# B&R Automation Studio project BoostTest
Automation Studio 6.7.2.9; technology packages: OpcUaCs 6.0.0

## Configuration CgAutomation

CPU X20EM0611, AutomationRuntime 6.3.4, Build 11.3.0, Vc 6.0.0

### Task classes (Cpu.sw)
```
Cyclic#1:
  Prg01 <- Machine.Prg01.prg
Cyclic#2:
  Prg02 <- Machine.Prg02.prg
Binaries: udbdef, FWRules, TCData, sysconf, iomap, ashwd, BRRole, asfw, arconfig, ashwac, UaCsConfig
Libraries: sys_lib, runtime, CFrw, CAlarm, astime, AsIecCon, CPrg01, CPrg02
```

### Hardware
```
X20EM0611 : X20EM0611 v1.1.1.0
  Connector IF2:
    ActivateDevice = 1
  ConfigurationID = BoostTest_CgAutomation
  Simulation = 1
  FileDevice1
  FileDeviceName1 = USER
  FileDevicePath1 = USER_PATH
```

### BRRole.brrole - X20EM0611/AccessAndSecurity/UserRoleSystem/BRRole.brrole
```
Element BR_Anonymous (Type=BRRole)
Element BR_Engineer (Type=BRRole)
Element BR_Observer (Type=BRRole)
Element BR_SafetyAdmin (Type=BRRole)
Element BR_SecurityAdmin (Type=BRRole)
```

- Safety project (password-protected, skipped)

## Logical view

Binary libraries used (declarations not repeated): operator, runtime, AsIecCon, astime, sys_lib

### Package Logical/Libraries - Global libraries

### Framework.st
```iecst
ACTION aFrwInit:
	ST_name(0, ADR(sObjName), 0);
END_ACTION

ACTION aFrwCyclic:

	aPreStateExt;
	aCallRessource;
	CASE stModuleData.enModuleState OF

		enState_Initialising:
            aInitialisingExt;
            IF (stModuleData.bInitDone) THEN
                stModuleData.enModuleState := enState_Stopped;
            END_IF

		enState_Stopped:
			aStoppedExt;

		enState_Running:
			aRunningExt;

		ELSE
			stModuleData.enModuleState := enState_Initialising;
	END_CASE

	aPostStateExt;

END_ACTION

ACTION aRessource_01:
    udiRessource_01 := udiRessource_01 + 1;
END_ACTION

ACTION aRessource_02:
    udiRessource_02 := udiRessource_02 + 2;
END_ACTION
```

### Framework.var
```iecst
VAR
    _ii : INT;
    sObjName : STRING[10];
    dstAlarm : REFERENCE TO tstCFrw_AlarmType;
END_VAR
(*Sub-States*)
VAR
    stInitialisingExt : tstInitialisingExt;
    stRunExt : tstRunExt;
    New_Variable : USINT;
END_VAR
```

### Library Logical/Framework/Ressources/CFrw (IEC)

#### Types.typ - Exported data types
```iecst
TYPE
	tenCFrw_States :
		(
		enState_Initialising,
		enState_Stopped,
		enState_Running
		);
	tstCFrw_AlarmType : 	STRUCT
		sDefaultText : STRING[255];
		udiCode : UDINT;
		uiSeverity : UINT;
	END_STRUCT;
END_TYPE
```

### Ressource_01.var
```iecst
VAR
    udiRessource_01 : UDINT;
END_VAR
```

### Ressource_01.st
```iecst
ACTION aCallRessource:
    aRessource_01;
    aReferencedAction;
END_ACTION

ACTION aReferencedAction:
    aLocalAction;
END_ACTION
```

### Ressource_02.var
```iecst
VAR
    udiRessource_02 : UDINT;
END_VAR
```

### Ressource_02.st
```iecst
ACTION aCallRessource:
    aRessource_02;
END_ACTION
```

### Program Logical/Framework/Template/Template (IEC)

- Framework.st (reference to Logical/Framework/Ressources/Framework.st)

- Framework.var (reference to Logical/Framework/Ressources/Framework.var)

#### Cyclic.st - Cyclic code
```iecst
PROGRAM _CYCLIC
	(* Insert code here *)
	 aFrwCyclic;
END_PROGRAM
```

#### Init.st - Init code
```iecst
PROGRAM _INIT
	(* Insert code here *)
	aFrwInit;

END_PROGRAM
```

#### Exit.st - Exit code
```iecst
PROGRAM _EXIT
	(* Insert code here *)

END_PROGRAM
```

#### Template.typ - Local data types
```iecst
TYPE
    tstAlarmList :     STRUCT
        stFrwAlarms : tstCAlarm_FrwAlarmListType;
        stModuleAlarms : tst_TEMPL_AlarmType;
    END_STRUCT;
    tst_TEMPL_AlarmType :     STRUCT
        stAlarm500000 : tstAlarm500000;
    END_STRUCT;
END_TYPE

(*States*)

TYPE
    tstInitialisingExt :     STRUCT
        enState : tenInitialisingExt;
    END_STRUCT;
    tenInitialisingExt :
        (
        enInitialisingExt_EntryAction,
        enInitialisingExt_, (*insert machine specific states here*)
        enInitialisingExt_Done
        );
    tstRunExt :     STRUCT
        enState : tenRunExt;
    END_STRUCT;
    tenRunExt :
        (
        enRunExt_EntryAction,
        enRunExt_, (*insert machine specific states here*)
        enRunExt_Done
        );
END_TYPE
```

#### Template.var - Local variables
```iecst
VAR
    stAlarmList : tstAlarmList;
    stModuleData : tstC_TEMPL_Data;
END_VAR
```

#### PreStateExt.st
```iecst
ACTION aPreStateExt:

END_ACTION
```

#### States.st
```iecst
ACTION aInitialisingExt:
    CASE stInitialisingExt.enState OF
        enInitialisingExt_EntryAction:
            stInitialisingExt.enState := enInitialisingExt_;
        enInitialisingExt_:
            (*implement machine specific code here*)
            stInitialisingExt.enState := enInitialisingExt_Done;
        enInitialisingExt_Done:
            (*set bInitDone := TRUE if initialising is completed*)
            stModuleData.bInitDone := TRUE;
        ELSE
            ;
    END_CASE
END_ACTION

ACTION aStoppedExt:

END_ACTION

ACTION aRunningExt:

END_ACTION
```

#### PostStateExt.st
```iecst
ACTION aPostStateExt:

END_ACTION
```

### Library Logical/Framework/Template/C_TEMPL_ (IEC)

#### C_TEMPL_.typ - Exported data types
```iecst
TYPE
    tstC_TEMPL_Data :     STRUCT
        enModuleState : tenCFrw_States;
        bInitDone : BOOL;
        stPar : tstC_TEMPL_Par;
    END_STRUCT;
    tstC_TEMPL_Par :     STRUCT
        udiPar01 : UDINT;
    END_STRUCT;
END_TYPE
```

### Library Logical/Machine/CAlarm (IEC)

#### Types.typ - Exported data types
```iecst
(*Framework*)

TYPE
	tstAlarm100000 :tstCFrw_AlarmType := (sDefaultText:='Message 100000',udiCode:=100000);
	tstAlarm100001 :tstCFrw_AlarmType := (sDefaultText:='Message 100001',udiCode:=100001);
	tstAlarm100002 :tstCFrw_AlarmType := (sDefaultText:='Message 100002',udiCode:=100002);
	tstCAlarm_FrwAlarmListType : 	STRUCT
		stAlarm100000 : tstAlarm100000;
		stAlarm100001 : tstAlarm100001;
		stAlarm100002 : tstAlarm100002;
	END_STRUCT;
END_TYPE

(*Process*)

TYPE
	tstAlarm500000 :tstCFrw_AlarmType := (sDefaultText:='Message 500000',udiCode:=500000);
	tstAlarm500001 :tstCFrw_AlarmType := (sDefaultText:='Message 500001',udiCode:=500001);
END_TYPE
```

### Program Logical/Machine/Prg01 (IEC)

- Framework.st (reference to Logical/Framework/Ressources/Framework.st)

- Framework.var (reference to Logical/Framework/Ressources/Framework.var)

- Ressource_01.var (reference to Logical/Framework/Ressources/Ressource_01/Ressource_01.var)

- Ressource_01.st (reference to Logical/Framework/Ressources/Ressource_01/Ressource_01.st)

#### Action.st
```iecst
ACTION aLocalAction:
    sText := 'aLocalAction called';
END_ACTION
```

#### Cyclic.st - Cyclic code
```iecst
PROGRAM _CYCLIC
	(* Insert code here *)
    aFrwCyclic;
    udiRessource_01;
END_PROGRAM
```

#### Init.st - Init code
```iecst
PROGRAM _INIT
	(* Insert code here *)
	aFrwInit;

END_PROGRAM
```

#### Exit.st - Exit code
```iecst
PROGRAM _EXIT
	(* Insert code here *)

END_PROGRAM
```

#### Prg01.typ - Local data types
```iecst
TYPE
    tstAlarmList :     STRUCT
        stFrwAlarms : tstCAlarm_FrwAlarmListType;
        stModuleAlarms : tstPrg01_AlarmType;
    END_STRUCT;
    tstPrg01_AlarmType :     STRUCT
        stAlarm500000 : tstAlarm500000;
    END_STRUCT;
END_TYPE

(*States*)

TYPE
    tstInitialisingExt :     STRUCT
        enState : tenInitialisingExt;
    END_STRUCT;
    tenInitialisingExt :
        (
        enInitialisingExt_EntryAction,
        enInitialisingExt_InitPrg01, (*insert machine specific states here*)
        enInitialisingExt_Done
        );
    tstRunExt :     STRUCT
        enState : tenRunExt;
    END_STRUCT;
    tenRunExt :
        (
        enRunExt_EntryAction,
        enRunExt_, (*insert machine specific states here*)
        enRunExt_Done
        );
    tstDebugStruct :     STRUCT
        bFlag : BOOL;
        diValue : DINT;
    END_STRUCT;
END_TYPE
```

#### Prg01.var - Local variables
```iecst
VAR
    stAlarmList : tstAlarmList;
    stModuleData : tstCPrg01Data;
    sText : STRING[80];
    pDebugArray : UDINT;
    astDebugArray : ARRAY[0..1] OF tstDebugStruct;
    dastDebugArray : REFERENCE TO ARRAY[0..1] OF tstDebugStruct;
END_VAR
```

#### PreStateExt.st
```iecst
ACTION aPreStateExt:
    pDebugArray := ADR(astDebugArray);
    dastDebugArray ACCESS pDebugArray;
END_ACTION
```

#### States.st
```iecst
ACTION aInitialisingExt:

    CASE stInitialisingExt.enState OF
        enInitialisingExt_EntryAction:
            stInitialisingExt.enState := enInitialisingExt_InitPrg01;
        enInitialisingExt_InitPrg01:
            (*implement machine specific code here*)
            stInitialisingExt.enState := enInitialisingExt_Done;
        enInitialisingExt_Done:
            (*set bInitDone := TRUE if initialising is completed*)
            stModuleData.bInitDone := TRUE;
        ELSE
            ;
    END_CASE
END_ACTION

ACTION aStoppedExt:

	FOR _ii := 0 TO 5 DO
		;
	END_FOR

END_ACTION

ACTION aRunningExt:

END_ACTION
```

#### PostStateExt.st
```iecst
ACTION aPostStateExt:

	FOR _ii := 0 TO (SIZEOF(stAlarmList.stFrwAlarms)/SIZEOF(dstAlarm) - 1) DO
		dstAlarm ACCESS ADR(stAlarmList.stFrwAlarms) + _ii * SIZEOF(dstAlarm);
	END_FOR

END_ACTION
```

### Library Logical/Machine/CPrg01 (IEC)

#### CPrg01.typ - Exported data types
```iecst
TYPE
    tstCPrg01Data :     STRUCT
        enModuleState : tenCFrw_States;
        bInitDone : BOOL;
        stPar : tstCPrg01Par;
    END_STRUCT;
    tstCPrg01Par :     STRUCT
        udiPar01 : UDINT;
    END_STRUCT;
END_TYPE
```

### Program Logical/Machine/Prg02 (IEC)

- Framework.st (reference to Logical/Framework/Ressources/Framework.st)

- Framework.var (reference to Logical/Framework/Ressources/Framework.var)

- Ressource_02.var (reference to Logical/Framework/Ressources/Ressource_02/Ressource_02.var)

- Ressource_02.st (reference to Logical/Framework/Ressources/Ressource_02/Ressource_02.st)

#### Cyclic.st - Cyclic code
```iecst
PROGRAM _CYCLIC
	(* Insert code here *)
    aFrwCyclic;
    udiRessource_02;
END_PROGRAM
```

#### Init.st - Init code
```iecst
PROGRAM _INIT
	(* Insert code here *)
	aFrwInit;

END_PROGRAM
```

#### Exit.st - Exit code
```iecst
PROGRAM _EXIT
	(* Insert code here *)

END_PROGRAM
```

#### Prg02.typ - Local data types
```iecst
TYPE
    tstAlarmList :     STRUCT
        stFrwAlarms : tstCAlarm_FrwAlarmListType;
        stModuleAlarms : tstPrg02_AlarmType;
    END_STRUCT;
    tstPrg02_AlarmType :     STRUCT
        stAlarm500001 : tstAlarm500001;
    END_STRUCT;
END_TYPE

(*States*)

TYPE
    tstInitialisingExt :     STRUCT
        enState : tenInitialisingExt;
    END_STRUCT;
    tenInitialisingExt :
        (
        enInitialisingExt_EntryAction,
        enInitialisingExt_InitPrg02, (*insert machine specific states here*)
        enInitialisingExt_Done
        );
    tstRunExt :     STRUCT
        enState : tenRunExt;
    END_STRUCT;
    tenRunExt :
        (
        enRunExt_EntryAction,
        enRunExt_, (*insert machine specific states here*)
        enRunExt_Done
        );
END_TYPE
```

#### Prg02.var - Local variables
```iecst
VAR
    stAlarmList : tstAlarmList;
    stModuleData : tstCPrg02Data;
    uiVariable : UINT;
END_VAR
```

#### PreStateExt.st
```iecst
ACTION aPreStateExt:

END_ACTION
```

#### States.st
```iecst
ACTION aInitialisingExt:
    CASE stInitialisingExt.enState OF
        enInitialisingExt_EntryAction:
            stInitialisingExt.enState := enInitialisingExt_InitPrg02;
        enInitialisingExt_InitPrg02:
            stInitialisingExt.enState := enInitialisingExt_Done;
        enInitialisingExt_Done:
            (*set bInitDone := TRUE if initialising is completed*)
            stModuleData.bInitDone := TRUE;
        ELSE
            ;
    END_CASE
END_ACTION

ACTION aStoppedExt:

	FOR _ii := 0 TO 5 DO
		;
	END_FOR
	uiVariable;
    fTestBitset(ADR(uiVariable));

END_ACTION

ACTION aRunningExt:

END_ACTION
```

#### PostStateExt.st
```iecst
ACTION aPostStateExt:

	stAlarmList;
END_ACTION
```

### Library Logical/Machine/CPrg02 (IEC)

#### CPrg02.typ - Exported data types
```iecst
TYPE
    tstCPrg02Data :     STRUCT
        enModuleState : tenCFrw_States;
        bInitDone : BOOL;
        stPar : tstCPrg02Par;
    END_STRUCT;
    tstCPrg02Par :     STRUCT
        udiPar01 : UDINT;
    END_STRUCT;
END_TYPE
```

#### CPrg02.fun - Exported functions and function blocks
```iecst
{REDUND_ERROR} FUNCTION fTestBitset : BOOL (*TODO: Add your comment here*) (*$GROUP=User,$CAT=User,$GROUPICON=User.png,$CATICON=User.png*)
    VAR_INPUT
        i_uiBitset : REFERENCE TO UINT;
    END_VAR
END_FUNCTION
```

#### fTestBitset.st
```iecst
(* TODO: Add your comment here *)
FUNCTION fTestBitset
    fTestBitset := TRUE;

    i_uiBitset.0 := TRUE;
    i_uiBitset.1 := FALSE;

    // Nur für Boost-Demo:
    fTestBitset := fTestBitset AND TRUE;
END_FUNCTION
```
